(* IEC 61131-3 sources: Elmo_Master/Lasal_PRG/Welcon8Axis_EtherCAT_Test_With_RobotAxis/Network, 1 file *)

(* ---- ConfigObjects.st ---- *)
FUNCTION GLOBAL TAB TASK_CONF
_K_TASK, _K_REAL,
_K_END_VAR,

_K_TASK, _K_CYCLIC,
_K_END_VAR,

_K_TASK, _K_BACKGROUND,
_K_END_VAR,

_K_END_CONF
END_FUNCTION

FUNCTION GLOBAL TAB IPR_CONF
_K_IPR
	0$UINT,
_K_END_VAR,
_K_END_CONF
END_FUNCTION

FUNCTION GLOBAL TAB CONFIG_TABLES
00115$UINT,
0$UINT, 1, 58, "_AXISBASE",
0$UINT, 0, 5, "_CAN",
0$UINT, 1, 11, "_CANLIB",
0$UINT, 1, 0, "_CHECKSUM",
0$UINT, 1, 20, "_FILESYS",
0$UINT, 0, 5, "_LINKER",
0$UINT, 1, 0, "_LMCABSENCODER",
0$UINT, 1, 120, "_LMCAXIS",
0$UINT, 2, 111, "_LMCAXISBASE",
0$UINT, 1, 32, "_LMCAXISREF",
0$UINT, 1, 42, "_LMCAXISVIS",
0$UINT, 1, 63, "_LMCAXISVISINT",
0$UINT, 1, 0, "_LMCAXISVISLOGHANDLE",
0$UINT, 1, 0, "_LMCAXISVISLOGVIEWER",
0$UINT, 1, 13, "_LMCAXISVISPARA",
0$UINT, 1, 2, "_LMCAXISVOVMONITORING",
0$UINT, 1, 18, "_LMCBASECOORD",
0$UINT, 1, 7, "_LMCBELTAXIS",
0$UINT, 1, 5, "_LMCCALCMODELBASE",
0$UINT, 1, 2, "_LMCCALCMODELCONTROLLER",
0$UINT, 1, 24, "_LMCMATH_SO3",
0$UINT, 1, 75, "_LMCMATHFUNCTIONS",
0$UINT, 1, 1, "_LMCMODULEBASE",
0$UINT, 3, 0, "_LMCPROFILE",
0$UINT, 4, 0, "_LMCPROFILEBASE",
0$UINT, 1, 53, "_LMCPROFILEBUFFER",
0$UINT, 1, 44, "_LMCPROFILELOG",
0$UINT, 1, 30, "_LMCPROFILEVIS",
0$UINT, 1, 20, "_LMCPROFILEVISAXIS",
0$UINT, 1, 41, "_LMCPROFILEVISINT",
0$UINT, 1, 30, "_LMCPROFILEVISMOVEPARA",
0$UINT, 1, 0, "_LMCPUBLISHER",
0$UINT, 1, 11, "_LMCREFBASE",
0$UINT, 2, 22, "_LMCROBOTBASE",
0$UINT, 1, 42, "_LMCROBOTLOG",
0$UINT, 1, 21, "_LMCSAFETY",
0$UINT, 1, 2, "_LMCSPLINEBUFFER",
0$UINT, 1, 23, "_LMCTABLEBUFFER",
0$UINT, 1, 3, "_LMCTOOL",
0$UINT, 1, 1, "_MULTITASK",
0$UINT, 0, 5, "_OSKERNEL",
0$UINT, 1, 36, "_SERLIB",
0$UINT, 1, 1, "_SIGTCPCOMRECEIVE",
0$UINT, 1, 1, "_SIGTCPDATAMANAGER",
0$UINT, 2, 0, "_STDLIB",
0$UINT, 1, 4, "_SYNCMEASURE",
0$UINT, 1, 3, "_SYNCMEASUREECAT",
0$UINT, 1, 1, "_TASKOBJECTCONTROL",
0$UINT, 1, 2, "_UDPTRANSCEIVER",
0$UINT, 1, 3, "_UDPTRANSCEIVERINTERFACE",
0$UINT, 1, 21, "ASCII_BIN",
0$UINT, 2, 2, "BUSINTERFACESDIASINTERNAL",
0$UINT, 1, 47, "CONTROLLER",
0$UINT, 1, 1, "CP313_IOS",
0$UINT, 0, 4, "CRITICALSECTION",
0$UINT, 1, 1, "DATAMANAGER",
0$UINT, 1, 1, "DATAMANAGERFIFO",
0$UINT, 1, 0, "DATAMANAGERPRIORITY",
0$UINT, 2, 34, "DIASMASTER",
0$UINT, 1, 84, "DIASMASTERC",
0$UINT, 2, 26, "DIASMASTERMAIN",
0$UINT, 1, 1, "DIASMASTERPOSTSCAN",
0$UINT, 1, 3, "DRIVEAXISDS402",
0$UINT, 1, 0, "DRIVEAXISDS402_BASE",
0$UINT, 1, 2, "ECAT_DS402BASE",
0$UINT, 2, 3, "ECAT_MASTER_BASE",
0$UINT, 2, 1, "ECAT_SLAVE_BASE",
0$UINT, 1, 12, "EEPROM",
0$UINT, 1, 2, "ETHERCAT_HUB_BASE",
0$UINT, 2, 2, "ETHERCAT_PLC",
0$UINT, 1, 5, "GETCILINTERFACE",
0$UINT, 0, 2, "GETTASKHANDLE",
0$UINT, 1, 22, "HUB_BASE",
0$UINT, 2, 12, "HUB_BASE_ROOT",
0$UINT, 2, 37, "HWBASE",
0$UINT, 2, 57, "HWBASECDIAS",
0$UINT, 1, 1, "HWCLOGGING",
0$UINT, 6, 0, "HWCONTROL",
0$UINT, 1, 11, "HWCONTROLBASE",
0$UINT, 1, 1, "HWRTPOSTSCAN",
0$UINT, 1, 7, "I2CCDIAS",
0$UINT, 1, 0, "MERKER",
0$UINT, 1, 22, "MERKEREX",
0$UINT, 1, 0, "MOVESPLINETABLE",
0$UINT, 2, 77, "POSCONTROLLER",
0$UINT, 1, 9, "RAMFILE",
0$UINT, 1, 1, "RAMRINGBUFFER",
0$UINT, 0, 0, "ROBOT_HANDLER",
0$UINT, 3, 20, "SAFETYCDIAS_BASE",
0$UINT, 3, 0, "SAFETYMANAGER",
0$UINT, 1, 0, "SAFETYROUTINGTABLES",
0$UINT, 1, 5, "SAFETYUDP",
0$UINT, 2, 0, "SDIASBASE",
0$UINT, 1, 11, "SDIASHUBBASE",
0$UINT, 1, 100, "SDIASMANAGER",
0$UINT, 2, 8, "SDIASPLC",
0$UINT, 0, 46, "SIGCLIB",
0$UINT, 1, 11, "STRING",
0$UINT, 1, 86, "STRINGINTERNAL",
0$UINT, 1, 22, "SYNCCALL",
0$UINT, 0, 0, "TCP_MOTIONIF_DUMMY",
0$UINT, 1, 20, "TCPCOMMUNICATION",
0$UINT, 1, 0, "TCPCOMMUNICATIONLOGFILTER",
0$UINT, 0, 0, "UDPTRANSMISSION",
0$UINT, 2, 22, "VARAN_BASE",
0$UINT, 3, 9, "VARANMANAGER",
0$UINT, 2, 8, "VARANMANAGER_1",
0$UINT, 1, 27, "VARANMANAGER_BASE",
0$UINT, 1, 3, "VIRTUALBASEINIT",
0$UINT, 2, 12, "WATCHDOGDIAS",
0$UINT, 0, 0, "WELCON_1",
0$UINT, 0, 0, "WELCON_2",
0$UINT, 0, 0, "WELCON_3",
0$UINT, 0, 0, "WELCON_4",
0$UINT, 1, 4, "XXXBASE_IOS",
ONE_CFG$UINT, 0, 0, "ONE_Axis1",
ONE_CFG$UINT, 0, 0, "ONE_Axis2",
ONE_CFG$UINT, 0, 0, "ONE_Axis3",
ONE_CFG$UINT, 0, 0, "ONE_Axis4",
ONE_CFG$UINT, 0, 0, "ONE_Axis5",
ONE_CFG$UINT, 0, 0, "ONE_Axis6",
ONE_CFG$UINT, 0, 0, "ONE_Axis7",
ONE_CFG$UINT, 0, 0, "ONE_Axis8",
ONE_CFG$UINT, 0, 0, "ONE_DS402_Network",
ONE_CFG$UINT, 0, 0, "ONE_HW_Network",
ONE_CFG$UINT, 0, 0, "ONE_Robot_Network",
ONE_CFG$UINT, 0, 0, "ONE_TCPComNet",
ONE_CFG$UINT, 0, 0, "ONE_UDPComNet",
TASK_CFG$UINT, 0, 0, "TASK_CONF",
IPR_CFG$UINT, 0, 0, "IPR_CONF",
PRJ_CFG$UINT, 0, 0, "Welcon8Axis_EtherCAT_Test_With_RobotAxis",
END_FUNCTION

#ifdef __LSLLDR_IOELEMENTS__
FUNCTION GLOBAL TAB _IO_ELEMENTS_TAB
0001$UINT, 0001$UINT,
"**IOCONN_EMPTY**", "WELCON_11.RxPDO9_Controlword2",
0081$UINT,
"**IOCONN_EMPTY**", "DriveAxisDS402_Axis2.CiA_ControlWord",
"**IOCONN_EMPTY**", "DriveAxisDS402_Axis2.CiA_StatusWord",
"**IOCONN_EMPTY**", "DriveAxisDS402_Axis2.ModesOfOperation",
"**IOCONN_EMPTY**", "DriveAxisDS402_Axis2.ModesOfOperationDisplay",
"**IOCONN_EMPTY**", "DriveAxisDS402_Axis2.PositionActualValue",
"**IOCONN_EMPTY**", "DriveAxisDS402_Axis2.TargetPosition",
"**IOCONN_EMPTY**", "DriveAxisDS402_Axis2.TargetTorque",
"**IOCONN_EMPTY**", "DriveAxisDS402_Axis2.TargetVelocity",
"**IOCONN_EMPTY**", "DriveAxisDS402_Axis2.TorqueActualValue",
"**IOCONN_EMPTY**", "DriveAxisDS402_Axis2.VelocityActualValue",
"**IOCONN_EMPTY**", "DriveAxisDS402_Axis2.Online",
"**IOCONN_EMPTY**", "DriveAxisDS402_Axis4.CiA_ControlWord",
"**IOCONN_EMPTY**", "DriveAxisDS402_Axis4.CiA_StatusWord",
"**IOCONN_EMPTY**", "DriveAxisDS402_Axis4.ModesOfOperation",
"**IOCONN_EMPTY**", "DriveAxisDS402_Axis4.ModesOfOperationDisplay",
"**IOCONN_EMPTY**", "DriveAxisDS402_Axis4.PositionActualValue",
"**IOCONN_EMPTY**", "DriveAxisDS402_Axis4.TargetPosition",
"**IOCONN_EMPTY**", "DriveAxisDS402_Axis4.TargetTorque",
"**IOCONN_EMPTY**", "DriveAxisDS402_Axis4.TargetVelocity",
"**IOCONN_EMPTY**", "DriveAxisDS402_Axis4.TorqueActualValue",
"**IOCONN_EMPTY**", "DriveAxisDS402_Axis4.VelocityActualValue",
"**IOCONN_EMPTY**", "DriveAxisDS402_Axis4.Online",
"**IOCONN_EMPTY**", "DriveAxisDS402_Axis8.CiA_ControlWord",
"**IOCONN_EMPTY**", "DriveAxisDS402_Axis8.CiA_StatusWord",
"**IOCONN_EMPTY**", "DriveAxisDS402_Axis8.ModesOfOperation",
"**IOCONN_EMPTY**", "DriveAxisDS402_Axis8.ModesOfOperationDisplay",
"**IOCONN_EMPTY**", "DriveAxisDS402_Axis8.PositionActualValue",
"**IOCONN_EMPTY**", "DriveAxisDS402_Axis8.TargetPosition",
"**IOCONN_EMPTY**", "DriveAxisDS402_Axis8.TargetTorque",
"**IOCONN_EMPTY**", "DriveAxisDS402_Axis8.TargetVelocity",
"**IOCONN_EMPTY**", "DriveAxisDS402_Axis8.TorqueActualValue",
"**IOCONN_EMPTY**", "DriveAxisDS402_Axis8.VelocityActualValue",
"**IOCONN_EMPTY**", "DriveAxisDS402_Axis8.Online",
"**IOCONN_EMPTY**", "PosController_Axis1.iHWErrors",
"**IOCONN_EMPTY**", "PosController_Axis1.oActive",
"**IOCONN_EMPTY**", "DriveAxisDS402_Axis6.CiA_ControlWord",
"**IOCONN_EMPTY**", "DriveAxisDS402_Axis6.CiA_StatusWord",
"**IOCONN_EMPTY**", "DriveAxisDS402_Axis6.ModesOfOperation",
"**IOCONN_EMPTY**", "DriveAxisDS402_Axis6.ModesOfOperationDisplay",
"**IOCONN_EMPTY**", "DriveAxisDS402_Axis6.PositionActualValue",
"**IOCONN_EMPTY**", "DriveAxisDS402_Axis6.TargetPosition",
"**IOCONN_EMPTY**", "DriveAxisDS402_Axis6.TargetVelocity",
"**IOCONN_EMPTY**", "DriveAxisDS402_Axis6.TargetTorque",
"**IOCONN_EMPTY**", "DriveAxisDS402_Axis6.TorqueActualValue",
"**IOCONN_EMPTY**", "DriveAxisDS402_Axis6.VelocityActualValue",
"**IOCONN_EMPTY**", "DriveAxisDS402_Axis6.Online",
"**IOCONN_EMPTY**", "PosController_Axis1.oOutputSignal",
"**IOCONN_EMPTY**", "PosController_Axis1.DriveEnabled",
"**IOCONN_EMPTY**", "PosController_Axis1.HWErrorQuit",
"**IOCONN_EMPTY**", "_LMCAxis_Axis1.ActPosition",
"**IOCONN_EMPTY**", "_LMCAxis_Axis1.HWReady",
"**IOCONN_EMPTY**", "_LMCAxis_Axis1.HWError",
"**IOCONN_EMPTY**", "_LMCAxis_Axis2.HWReady",
"**IOCONN_EMPTY**", "PosController_Axis3.iHWErrors",
"**IOCONN_EMPTY**", "PosController_Axis3.oActive",
"**IOCONN_EMPTY**", "PosController_Axis3.oOutputSignal",
"**IOCONN_EMPTY**", "PosController_Axis3.DriveEnabled",
"**IOCONN_EMPTY**", "PosController_Axis3.HWErrorQuit",
"**IOCONN_EMPTY**", "_LMCAxis_Axis3.HWReady",
"**IOCONN_EMPTY**", "_LMCAxis_Axis3.HWError",
"**IOCONN_EMPTY**", "_LMCAxis_Axis3.ActPosition",
"**IOCONN_EMPTY**", "PosController_Axis4.iHWErrors",
"**IOCONN_EMPTY**", "_LMCAxis_Axis4.HWReady",
"**IOCONN_EMPTY**", "PosController_Axis5.iHWErrors",
"**IOCONN_EMPTY**", "PosController_Axis5.oActive",
"**IOCONN_EMPTY**", "PosController_Axis5.oOutputSignal",
"**IOCONN_EMPTY**", "PosController_Axis5.DriveEnabled",
"**IOCONN_EMPTY**", "PosController_Axis5.HWErrorQuit",
"**IOCONN_EMPTY**", "_LMCAxis_Axis5.ActPosition",
"**IOCONN_EMPTY**", "_LMCAxis_Axis5.HWReady",
"**IOCONN_EMPTY**", "_LMCAxis_Axis5.HWError",
"**IOCONN_EMPTY**", "_LMCAxis_Axis6.HWReady",
"**IOCONN_EMPTY**", "PosController_Axis7.iHWErrors",
"**IOCONN_EMPTY**", "PosController_Axis7.oActive",
"**IOCONN_EMPTY**", "PosController_Axis7.oOutputSignal",
"**IOCONN_EMPTY**", "PosController_Axis7.DriveEnabled",
"**IOCONN_EMPTY**", "PosController_Axis7.HWErrorQuit",
"**IOCONN_EMPTY**", "_LMCAxis_Axis7.ActPosition",
"**IOCONN_EMPTY**", "_LMCAxis_Axis7.HWError",
"**IOCONN_EMPTY**", "_LMCAxis_Axis7.HWReady",
"**IOCONN_EMPTY**", "_LMCAxis_Axis8.HWReady",
END_FUNCTION
#endif //__LSLLDR_IOELEMENTS__

FUNCTION GLOBAL TAB CH_REDIRECT_EMB_TAB
0000$UINT,
00019$UINT,
"ECAT_DS402BASE;DEVICENAME", "\DEVICENAMESTR.DATA",
"ECAT_DS402BASE;PRODUCTREVISION", "\PRODUCTREVSTR.DATA",
"ECAT_MASTER_BASE;SOFTWAREVERSION", "\STRSOFTWAREVERSION.DATA",
"ECAT_SLAVE_BASE;DEVICENAME", "\DEVICENAMESTR.DATA",
"ECAT_SLAVE_BASE;PRODUCTREVISION", "\PRODUCTREVSTR.DATA",
"ETHERCAT_PLC;SOFTWAREVERSION", "\STRSOFTWAREVERSION.DATA",
"HWBASECDIAS;SERIALNO", "\SERIALNOSTR.DATA",
"SAFETYCDIAS_BASE;SERIALNO", "\SERIALNOSTR.DATA",
"SDIASBASE;SERIALNO", "\SERIALNOSTR.DATA",
"TCPCOMMUNICATION;TASKNAME", "\THREADNAME.DATA",
"VARAN_BASE;SERIALNO", "\SERIALNOSTR.DATA",
"WELCON_1;DEVICENAME", "\DEVICENAMESTR.DATA",
"WELCON_1;PRODUCTREVISION", "\PRODUCTREVSTR.DATA",
"WELCON_2;DEVICENAME", "\DEVICENAMESTR.DATA",
"WELCON_2;PRODUCTREVISION", "\PRODUCTREVSTR.DATA",
"WELCON_3;DEVICENAME", "\DEVICENAMESTR.DATA",
"WELCON_3;PRODUCTREVISION", "\PRODUCTREVSTR.DATA",
"WELCON_4;DEVICENAME", "\DEVICENAMESTR.DATA",
"WELCON_4;PRODUCTREVISION", "\PRODUCTREVSTR.DATA",
END_FUNCTION
